(* IEC 61131-3 sources: bcs-engineering-dsl/language/test/generating/functionblock_test/expected, 4 files *)

(* ---- SimpleLogicFB_decl.st ---- *)
FUNCTION_BLOCK SimpleLogicFB
VAR_INPUT
    iInput: BOOL;
    iInput2: INT;
END_VAR
VAR_OUTPUT
    oOutput: BOOL;
END_VAR
VAR
    iInputNegated: BOOL;
    R_TRIG_Instance1: R_TRIG;
    F_TRIG_Instance1: F_TRIG;
    TON_AfterInstance1: TON := (PT := T#1s);
    R_TRIG_AfterInstance1: R_TRIG;
END_VAR

(* ---- MAIN_decl.st ---- *)
PROGRAM MAIN
VAR
    TestFunctionBlock_input: BOOL := TRUE;
    TestFunctionBlock_input2: INT := 5;
    TestFunctionBlock_input3: BOOL := FALSE;
    TestFunctionBlock_input4: INT := 10;
    TestFunctionBlock_output: BOOL;
    TestFunctionBlock_output2: BOOL;
    SimpleLogicFBInstance1: SimpleLogicFB;
    SimpleLogicFBInstance2: SimpleLogicFB;
    F_TRIG_Instance3: F_TRIG;
END_VAR

(* ---- MAIN_impl.st ---- *)
// Control Unit 'TestFunctionBlock'
SimpleLogicFBInstance1(iInput:=TestFunctionBlock_input, iInput2:=TestFunctionBlock_input2);
TestFunctionBlock_output := SimpleLogicFBInstance1.oOutput;

SimpleLogicFBInstance2(iInput:=TestFunctionBlock_input3, iInput2:=TestFunctionBlock_input4);
TestFunctionBlock_output2 := SimpleLogicFBInstance2.oOutput;

F_TRIG_Instance3(CLK := TestFunctionBlock_input);
IF F_TRIG_Instance3.Q THEN
    TestFunctionBlock_output := FALSE;
END_IF;

(* ---- SimpleLogicFB_impl.st ---- *)
oOutput := iInput;
TON_AfterInstance1(IN := oOutput = TRUE);
R_TRIG_AfterInstance1(CLK := TON_AfterInstance1.Q);
IF R_TRIG_AfterInstance1.Q THEN
    oOutput := FALSE;
END_IF;
R_TRIG_Instance1(CLK := iInput);
IF R_TRIG_Instance1.Q THEN
    oOutput := TRUE;
END_IF;
F_TRIG_Instance1(CLK := iInput);
IF F_TRIG_Instance1.Q THEN
    oOutput := FALSE;
END_IF;
